Fanuc KAREL source: NM0041.KL

PROGRAM NM0041
%STACKSIZE=65535
%PRIORITY=65535
%NOLOCKGROUP
ROUTINE IDI(P1 : INTEGER) : INTEGER FROM NM0041
ROUTINE IDR(P1 : REAL) : REAL FROM NM0041
ROUTINE RTEST FROM NM0041
ROUTINE IDI
BEGIN
RETURN((P1 + 1))
END IDI
ROUTINE IDR
BEGIN
RETURN((P1 + 1.0))
END IDR
ROUTINE RTEST
VAR
L1 : STRING[8]
L2 : ARRAY[3] OF INTEGER
L3 : ARRAY[3] OF REAL
S1 : INTEGER
U2C_13 : INTEGER
S2 : REAL
U2C_15 : REAL
U2C_16 : BOOLEAN
BEGIN
S1=1
U2C_13=2
S2=2.5
U2C_15=3.5
U2C_16=TRUE
L1='A'
L2[1]=2
L3[1]=2.5
-- UNSAFE_SOURCE_IR line 30: CALL_RESULT IDI(S1)
END RTEST
BEGIN
RTEST
END NM0041
